(* PLC project probe.project, CODESYS CODESYS V3.5 SP17 Patch 3 *)
(* stored: creationDateTime 2026-10-20T03:54:26.8748154, modificationDateTime 1601-01-01T03:00:00 *)

FUNCTION_BLOCK FB_ProbeOop2
  VAR_INPUT
    xIn : BOOL;
  END_VAR
  VAR
    iState : INT;
  END_VAR

            iState := iState + 1;

          

ACTION ActClear:
                iState := 0;

              
END_ACTION

METHOD Reset : BOOL
  VAR_INPUT
    iTo : INT;
  END_VAR
                  iState := iTo;
Reset := TRUE;

                
END_METHOD

PROPERTY State : INT
GET
                    State := iState;

                  
END_GET
SET
                    iState := State;

                  
END_SET
END_PROPERTY
END_FUNCTION_BLOCK
